(* IEC 61131-3 sources: llm-plc-st-eval/data/processed_definitivo/gpt-4o-2024-08-06/A3/few_shot, 3 files *)

(* ---- ejec_1.st ---- *)
FUNCTION_BLOCK FB_Com
VAR_INPUT
    txReq : BOOL; (* Solicitud de transmision *)
    rxOk : BOOL; (* Confirmacion de recepcion *)
    rxData : INT; (* Datos recibidos *)
END_VAR
VAR_OUTPUT
    txData : INT; (* Datos a transmitir *)
    ocupado : BOOL; (* Indicador de intercambio en curso *)
    ok : BOOL; (* Indicador de exito *)
    error : BOOL; (* Indicador de error *)
    nIntentos : INT; (* Numero de intento actual *)
END_VAR
VAR
    txReqPrev : BOOL; (* Estado previo de txReq *)
    intentoActual : INT; (* Contador de intentos *)
    tTimeout : TON; (* Temporizador de timeout *)
    intercambioActivo : BOOL; (* Indicador de intercambio activo *)
END_VAR

(* Inicializacion de variables *)
IF NOT intercambioActivo THEN
    IF txReq AND NOT txReqPrev THEN
        (* Inicio de un nuevo intercambio *)
        txData := 100;
        ocupado := TRUE;
        ok := FALSE;
        error := FALSE;
        intentoActual := 1;
        nIntentos := intentoActual;
        intercambioActivo := TRUE;
        tTimeout(IN := TRUE, PT := T#500MS);
    END_IF
ELSE
    (* Proceso de intercambio en curso *)
    tTimeout(IN := NOT tTimeout.Q); (* Reiniciar temporizador si no ha expirado *)

    IF rxOk AND (rxData = txData) THEN
        (* Intento exitoso *)
        ok := TRUE;
        ocupado := FALSE;
        intercambioActivo := FALSE;
    ELSIF tTimeout.Q THEN
        (* Intento fallido, verificar siguiente intento *)
        intentoActual := intentoActual + 1;
        IF intentoActual > 3 THEN
            (* Todos los intentos fallaron *)
            error := TRUE;
            ocupado := FALSE;
            intercambioActivo := FALSE;
        ELSE
            (* Iniciar siguiente intento *)
            nIntentos := intentoActual;
            tTimeout(IN := TRUE, PT := T#500MS);
        END_IF
    END_IF
END_IF

(* Actualizar estado previo de txReq *)
txReqPrev := txReq;
END_FUNCTION_BLOCK

(* ---- ejec_2.st ---- *)
FUNCTION_BLOCK FB_Com
VAR_INPUT
    txReq : BOOL; (* Solicitud de transmisión *)
    rxOk : BOOL; (* Confirmación de recepción *)
    rxData : INT; (* Datos recibidos *)
END_VAR
VAR_OUTPUT
    txData : INT; (* Datos a transmitir *)
    ocupado : BOOL; (* Indica si el intercambio está en curso *)
    ok : BOOL; (* Indica si el intercambio fue exitoso *)
    error : BOOL; (* Indica si el intercambio falló *)
    nIntentos : INT; (* Número de intento actual *)
END_VAR
VAR
    intentoActual : INT := 0; (* Contador de intentos *)
    valorPrueba : INT := 100; (* Valor de prueba a transmitir *)
    tLimite : TON; (* Temporizador de límite de tiempo *)
    txReqAnt : BOOL := FALSE; (* Estado anterior de txReq *)
    intercambioEnCurso : BOOL := FALSE; (* Estado del intercambio *)
END_VAR

(* Detectar flanco ascendente de txReq *)
IF txReq AND NOT txReqAnt THEN
    IF NOT intercambioEnCurso THEN
        (* Iniciar nuevo intercambio *)
        txData := valorPrueba;
        ocupado := TRUE;
        ok := FALSE;
        error := FALSE;
        intentoActual := 1;
        intercambioEnCurso := TRUE;
        tLimite(IN := TRUE, PT := T#500MS);
    END_IF;
END_IF;

(* Control de intentos y recepción *)
IF intercambioEnCurso THEN
    IF tLimite.Q THEN
        (* Tiempo límite alcanzado, intento fallido *)
        intentoActual := intentoActual + 1;
        IF intentoActual > 3 THEN
            (* Todos los intentos fallaron *)
            error := TRUE;
            ocupado := FALSE;
            intercambioEnCurso := FALSE;
        ELSE
            (* Iniciar nuevo intento *)
            tLimite(IN := TRUE, PT := T#500MS);
        END_IF;
    ELSIF rxOk AND (rxData = valorPrueba) THEN
        (* Intento exitoso *)
        ok := TRUE;
        ocupado := FALSE;
        intercambioEnCurso := FALSE;
    END_IF;
END_IF;

(* Actualizar salidas *)
nIntentos := intentoActual;

(* Almacenar estado anterior de txReq *)
txReqAnt := txReq;
END_FUNCTION_BLOCK

(* ---- ejec_3.st ---- *)
FUNCTION_BLOCK FB_Com
VAR_INPUT
    txReq : BOOL; (* Solicitud de transmision *)
    rxOk : BOOL; (* Confirmacion de recepcion *)
    rxData : INT; (* Datos recibidos *)
END_VAR
VAR_OUTPUT
    txData : INT; (* Datos a transmitir *)
    ocupado : BOOL; (* Indicador de intercambio en curso *)
    ok : BOOL; (* Indicador de intercambio exitoso *)
    error : BOOL; (* Indicador de error en el intercambio *)
    nIntentos : INT; (* Numero de intento actual *)
END_VAR
VAR
    txReqPrev : BOOL; (* Estado previo de txReq *)
    intentoActual : INT; (* Contador de intentos *)
    tTimeout : TON; (* Temporizador de timeout *)
    intercambioActivo : BOOL; (* Indicador de intercambio activo *)
END_VAR

(* Inicializacion de variables *)
IF NOT intercambioActivo THEN
    IF txReq AND NOT txReqPrev THEN
        (* Inicio de un nuevo intercambio *)
        txData := 100;
        ocupado := TRUE;
        ok := FALSE;
        error := FALSE;
        intentoActual := 1;
        nIntentos := intentoActual;
        intercambioActivo := TRUE;
        tTimeout(IN := TRUE, PT := T#500MS);
    END_IF;
ELSE
    (* Proceso de intercambio en curso *)
    IF tTimeout.Q THEN
        (* Timeout del intento actual *)
        intentoActual := intentoActual + 1;
        IF intentoActual > 3 THEN
            (* Todos los intentos fallaron *)
            error := TRUE;
            ocupado := FALSE;
            intercambioActivo := FALSE;
        ELSE
            (* Iniciar siguiente intento *)
            nIntentos := intentoActual;
            tTimeout(IN := TRUE, PT := T#500MS);
        END_IF;
    ELSIF rxOk AND (rxData = txData) THEN
        (* Intento exitoso *)
        ok := TRUE;
        ocupado := FALSE;
        intercambioActivo := FALSE;
    END_IF;
END_IF;

(* Actualizar estado previo de txReq *)
txReqPrev := txReq;
END_FUNCTION_BLOCK
